TYPE "ST_StateFlag"
VERSION : 0.1
   STRUCT
      Key : String[120];
      Value : Bool;
      Since : LDT;
      Stale : Bool;
   END_STRUCT;

END_TYPE

